// TIA Portal project "session2" (V18)

(* hardware
DEVICE "S7-1200 station_1"  S7-1200 Station
   slot 0: "Rack_0"  S7-1200 Rack  Rack  V1.0
   slot 1: "PLC_1"  CPU 1215C DC/DC/DC  6ES7 215-1AG40-0XB0  V4.6
   slot 2: "SM 1278_1"  4SI IO link  6ES7 278-4BD32-0XB0  V2.1
   slot 3: "DI 2/DQ 2x24VDC_1"  DI2/DQ2 signal board  6ES7 223-0BD30-0XB0  V1.0
DEVICE "HMI_1"  KTP700 Basic PN
   slot 0: "HMI_1"  KTP700 Basic PN  6AV2 123-2GB03-0AX0  17.0.0.0
   slot 1: "HMI_RT_1"  KTP700 Basic PN  6AV2 123-2GB03-0AX0  17.0.0.0
   slot 5: "HMI_1.IE_CP_1"  PROFINET Interface  17.0.0.0
      slot 1: "PROFINET Interface_1"  PROFINET Interface
         slot 1: "Port_1"  Port
DEVICE "GSD device_1"  GSD.Device.PN
   slot 0: "Rack"  Rack  V1.0
   slot 0: "ur3ln"  V1.0  00000
      slot 0: "V1.0"  V1.0
      slot 1: "Interface"  Interface
         slot 1: "RJ45 10/100 MBit/s"  RJ45 10/100 MBit/s
   slot 5: "5_T2O General Purpose Bit Registers_1"  5_T2O General Purpose Bit Registers  1.0
      slot 0: "5_T2O General Purpose Bit Registers"  5_T2O General Purpose Bit Registers
   slot 9: "9_O2T General Purpose Registers 1_1"  9_O2T General Purpose Registers 1  1.0
      slot 0: "9_O2T General Purpose Registers 1"  9_O2T General Purpose Registers 1
*)

// ===== PLC "PLC_1"  CPU 1215C DC/DC/DC =====

VAR_GLOBAL   // PLC tag table "Default tag table"
   "x5" AT %I4.0 : Bool;
   "b1" AT %I1.3 : Bool;
   "b2" AT %I1.4 : Bool;
   "km1" AT %Q1.0 : Bool;
   "km2" AT %Q1.1 : Bool;
   "etap0" AT %M1.0 : Bool;
   "etap1" AT %M1.1 : Bool;
   "etap2" AT %M1.2 : Bool;
   "etap3" AT %M1.3 : Bool;
   "temps" AT %M10.0 : Bool;
   "pos int" AT %MW40 : Word;
   "loop" AT %M12.0 : Bool;
   "input compteur" AT %MW20 : Int;
   "output compteur" AT %MW80 : Int;
   "reset" AT %M5.1 : Bool;
   "Marche" AT %M5.0 : Bool;
   "Temps input" AT %MD30 : Time;
   "temps output" AT %MD34 : Time;
   "Off" AT %M5.2 : Bool;
   "Pos" AT %MW42 : Word;
   "Clock_Byte" AT %MB100 : Byte;
   "Clock_10Hz" AT %M100.0 : Bool;
   "Clock_5Hz" AT %M100.1 : Bool;
   "Clock_2.5Hz" AT %M100.2 : Bool;
   "Clock_2Hz" AT %M100.3 : Bool;
   "Clock_1.25Hz" AT %M100.4 : Bool;
   "Clock_1Hz" AT %M100.5 : Bool;
   "Clock_0.625Hz" AT %M100.6 : Bool;
   "Clock_0.5Hz" AT %M100.7 : Bool;
   "Courant Sig Aut" AT %IW64 : Int;
   "Courant NormX" AT %MD400 : Real;
   "Courant ScaleX" AT %MD500 : Real;
   "Tension Sig Aut" AT %IW66 : Int;
   "Tension NormX" AT %MD600 : Real;
   "Tension ScaleX" AT %MD700 : Real;
   "km4" AT %MW704 : Int;
   "Port Ultrason" AT %IW10 : Word;
   "SubDistance" AT %MW90 : Word;
   "hauteur" AT %MW92 : Word;
   "Distance Manu" AT %MW94 : Word;
   "Nbr Pieces" AT %MW96 : Word;
   "INC" AT %I1.5 : Bool;
   "pos RFID" AT %MW46 : Word;
   "Puc_Data" AT %MW48 : Word;
   "Vitesse" AT %MW110 : Word;
   "Tag_1" AT %QW1000 : Word;
   "Valid" AT %Q150.0 : Bool;
   "Finish" AT %I150.0 : Bool;
   "Err" AT %MW2 : Int;
END_VAR

VAR_GLOBAL   // PLC tag table "RFID_table"
   "RFID_commandBteOut" AT %QB10 : Byte;
   "RFID_CmdStart" AT %Q11.0 : Bool;
   "RFID_CmdDesactivateAntenna" AT %Q11.3 : Bool;
   "RFID_Write_Data1" AT %QW12 : Word;
   "RFID_CommandByteIn" AT %IB10 : Byte;
   "RFID_CmdStartAcknowledge" AT %I11.0 : Bool;
   "RFID_CmdEnd" AT %I11.1 : Bool;
   "RFID_Tag Present" AT %I11.2 : Bool;
   "RFID_Antenna Deactivated" AT %I11.3 : Bool;
   "RFID_Read_Data 1" AT %IW12 : Word;
   "RFID Read_Data2" AT %IW14 : Word;
   "RFID_Read_Data 3" AT %IW16 : Word;
   "RFID_Read_Data4" AT %IW18 : Word;
END_VAR

VAR_GLOBAL   // PLC tag table "Web"
   "Web_CMD_StartMarche" AT %M0.0 : Bool;
   "Web_CMD_StopMarche" AT %M0.1 : Bool;
   "Web_CMD_Reset" AT %M0.2 : Bool;
END_VAR

DATA_BLOCK "Ultrason"   // DB2
{ S7_Optimized_Access := 'TRUE' }
VERSION : 0.1
   VAR
      Distance : Int;
      Hauteur : Int;
      "Nbr Voiture" : Int;
      "Distance 0" : Int := 300;
      inter : Int;
   END_VAR
BEGIN
END_DATA_BLOCK

DATA_BLOCK "Energy Meter"   // DB6
{ S7_Optimized_Access := 'TRUE' }
VERSION : 0.1
   VAR
      Parameter_connexion : TCON_IP_v4;
   END_VAR
BEGIN
   Parameter_connexion.InterfaceId := 64;
   Parameter_connexion.ID := 1;
   Parameter_connexion.ActiveEstablished := true;
   Parameter_connexion.RemoteAddress.ADDR[1] := 172;
   Parameter_connexion.RemoteAddress.ADDR[2] := 28;
   Parameter_connexion.RemoteAddress.ADDR[3] := 111;
   Parameter_connexion.RemoteAddress.ADDR[4] := 56;
   Parameter_connexion.RemotePort := 502;
END_DATA_BLOCK

DATA_BLOCK "node_red"   // DB9
{ S7_Optimized_Access := 'FALSE' }
VERSION : 0.1
   VAR
      courant : Real;
      tension : Real;
   END_VAR
BEGIN
END_DATA_BLOCK

// folder: System blocks/Program resources

DATA_BLOCK "IEC_Timer_0_DB"   // DB1
{ S7_Optimized_Access := 'TRUE' }
AUTHOR : Simatic
FAMILY : IEC
NAME : IEC_TMR
VERSION : 1.0
// stored: InstanceOfName IEC_TIMER
"IEC_TIMER"
BEGIN
END_DATA_BLOCK

DATA_BLOCK "IEC_Counter_0_DB_1"   // DB3
{ S7_Optimized_Access := 'TRUE' }
AUTHOR : Simatic
FAMILY : IEC
NAME : CNTR
VERSION : 1.0
// stored: InstanceOfName IEC_COUNTER
"IEC_COUNTER"
BEGIN
END_DATA_BLOCK

DATA_BLOCK "IEC_Counter_0_DB_2"   // DB4
{ S7_Optimized_Access := 'TRUE' }
AUTHOR : Simatic
FAMILY : IEC
NAME : CNTR
VERSION : 1.0
// stored: InstanceOfName IEC_COUNTER
"IEC_COUNTER"
BEGIN
END_DATA_BLOCK

DATA_BLOCK "IEC_Counter_0_DB"   // DB7
{ S7_Optimized_Access := 'TRUE' }
AUTHOR : Simatic
FAMILY : IEC
NAME : CNTR
VERSION : 1.0
// stored: InstanceOfName IEC_COUNTER
"IEC_COUNTER"
BEGIN
END_DATA_BLOCK

// folder: (top level)

FUNCTION "configurer" : Void   // FC1, LAD
{ S7_Optimized_Access := 'TRUE' }
VERSION : 0.1
BEGIN

REGION Network 1
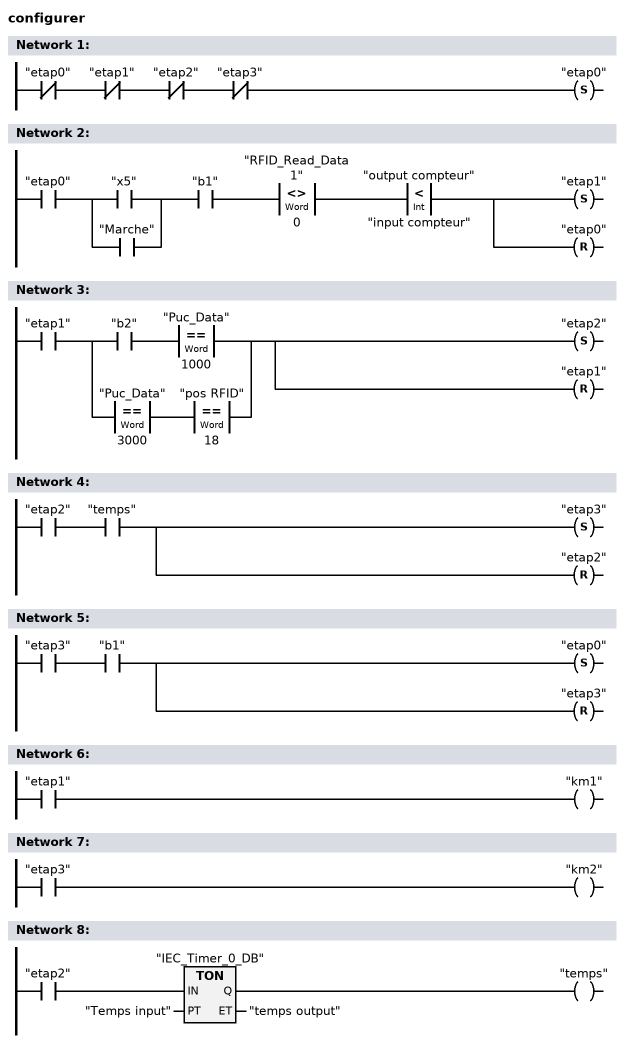
   RUNG wire#powerrail
      I_Contact( "etap0" )
      I_Contact( "etap1" )
      I_Contact( "etap2" )
      I_Contact( "etap3" )
      S_Coil( "etap0" )
   END_RUNG
   // the same network as SCL:
   IF NOT "etap0" AND NOT "etap1" AND NOT "etap2" AND NOT "etap3" THEN "etap0" := TRUE; END_IF;
END_REGION

REGION Network 2
   RUNG wire#powerrail
      Contact( "etap0" )
      wire#w1
      Contact( "x5" )
      wire#w2
      Contact( "b1" )
      { S7_Templates := "SrcType := Word" } NE_Contact(in1 := "RFID_Read_Data 1", in2 := 0)
      { S7_Templates := "SrcType := Int" } LT_Contact(in1 := "output compteur", in2 := "input compteur")
      wire#w3
      S_Coil( "etap1" )
   END_RUNG
   RUNG wire#w1
      Contact( "Marche" )
   END_RUNG wire#w2
   RUNG wire#w3
      R_Coil( "etap0" )
   END_RUNG
   // the same network as SCL:
   IF "etap0" AND ("x5" OR "Marche") AND "b1" AND ("RFID_Read_Data 1" <> 0) AND ("output compteur" < "input compteur") THEN
       "etap1" := TRUE;
       "etap0" := FALSE;
   END_IF;
END_REGION

REGION Network 3
   RUNG wire#powerrail
      Contact( "etap1" )
      wire#w1
      Contact( "b2" )
      { S7_Templates := "SrcType := Word" } EQ_Contact(in1 := "Puc_Data", in2 := 1000)
      wire#w2
      S_Coil( "etap2" )
   END_RUNG
   RUNG wire#w1
      { S7_Templates := "SrcType := Word" } EQ_Contact(in1 := "Puc_Data", in2 := 3000)
      { S7_Templates := "SrcType := Word" } EQ_Contact(in1 := "pos RFID", in2 := 18)
   END_RUNG wire#w2
   RUNG wire#w2
      R_Coil( "etap1" )
   END_RUNG
   // the same network as SCL:
   IF "etap1" AND (("b2" AND ("Puc_Data" = 1000)) OR (("Puc_Data" = 3000) AND ("pos RFID" = 18))) THEN
       "etap2" := TRUE;
       "etap1" := FALSE;
   END_IF;
END_REGION

REGION Network 4
   RUNG wire#powerrail
      Contact( "etap2" )
      Contact( "temps" )
      wire#w1
      S_Coil( "etap3" )
   END_RUNG
   RUNG wire#w1
      R_Coil( "etap2" )
   END_RUNG
   // the same network as SCL:
   IF "etap2" AND "temps" THEN
       "etap3" := TRUE;
       "etap2" := FALSE;
   END_IF;
END_REGION

REGION Network 5
   RUNG wire#powerrail
      Contact( "etap3" )
      Contact( "b1" )
      wire#w1
      S_Coil( "etap0" )
   END_RUNG
   RUNG wire#w1
      R_Coil( "etap3" )
   END_RUNG
   // the same network as SCL:
   IF "etap3" AND "b1" THEN
       "etap0" := TRUE;
       "etap3" := FALSE;
   END_IF;
END_REGION

REGION Network 6
   RUNG wire#powerrail
      Contact( "etap1" )
      Coil( "km1" )
   END_RUNG
   // the same network as SCL:
   "km1" := "etap1";
END_REGION

REGION Network 7
   RUNG wire#powerrail
      Contact( "etap3" )
      Coil( "km2" )
   END_RUNG
   // the same network as SCL:
   "km2" := "etap3";
END_REGION

REGION Network 8
   "IEC_Timer_0_DB".TON(IN := "etap2", PT := "Temps input", ET => "temps output");
   "temps" := "IEC_Timer_0_DB".Q;
END_REGION
END_FUNCTION

FUNCTION "Conversion" : Void   // FC2, LAD
{ S7_Optimized_Access := 'TRUE' }
VERSION : 0.1
BEGIN

REGION Network 1
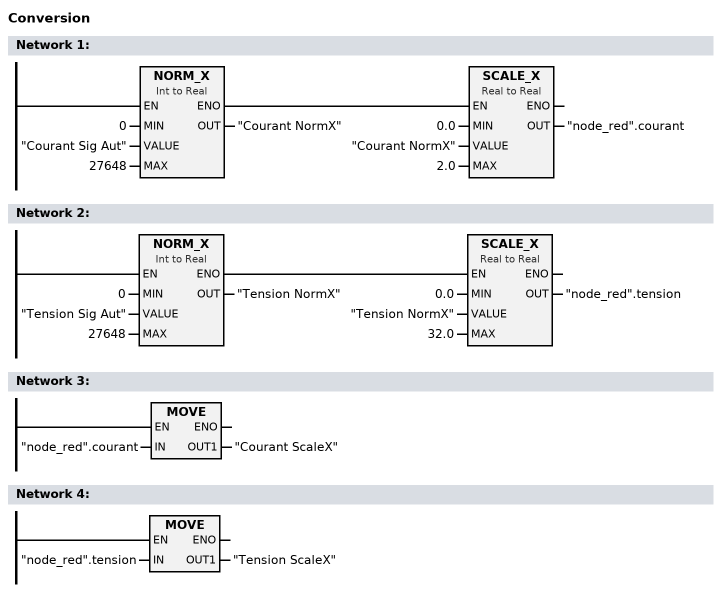
   RUNG wire#powerrail
      { S7_Templates := "[SrcType := Int, DestType := Real]" } Normalize(min := 0, value := "Courant Sig Aut", max := 27648, out => "Courant NormX")
      { S7_Templates := "[SrcType := Real, DestType := Real]" } Scale(min := 0.0, value := "Courant NormX", max := 2.0, out => "node_red".courant)
   END_RUNG
   // the same network as SCL:
   "Courant NormX" := NORM_X(MIN := 0, VALUE := "Courant Sig Aut", MAX := 27648);
   "node_red".courant := SCALE_X(MIN := 0.0, VALUE := "Courant NormX", MAX := 2.0);
END_REGION

REGION Network 2
   RUNG wire#powerrail
      { S7_Templates := "[SrcType := Int, DestType := Real]" } Normalize(min := 0, value := "Tension Sig Aut", max := 27648, out => "Tension NormX")
      { S7_Templates := "[SrcType := Real, DestType := Real]" } Scale(min := 0.0, value := "Tension NormX", max := 32.0, out => "node_red".tension)
   END_RUNG
   // the same network as SCL:
   "Tension NormX" := NORM_X(MIN := 0, VALUE := "Tension Sig Aut", MAX := 27648);
   "node_red".tension := SCALE_X(MIN := 0.0, VALUE := "Tension NormX", MAX := 32.0);
END_REGION

REGION Network 3
   RUNG wire#powerrail
      Move(in := "node_red".courant, out1 => "Courant ScaleX")
   END_RUNG
   // the same network as SCL:
   "Courant ScaleX" := "node_red".courant;
END_REGION

REGION Network 4
   RUNG wire#powerrail
      Move(in := "node_red".tension, out1 => "Tension ScaleX")
   END_RUNG
   // the same network as SCL:
   "Tension ScaleX" := "node_red".tension;
END_REGION
END_FUNCTION

FUNCTION "Ultrason Configuration" : Void   // FC3, LAD
{ S7_Optimized_Access := 'TRUE' }
VERSION : 0.1
   VAR_TEMP
      "inter 1" : Int;
   END_VAR
BEGIN

REGION Network 1
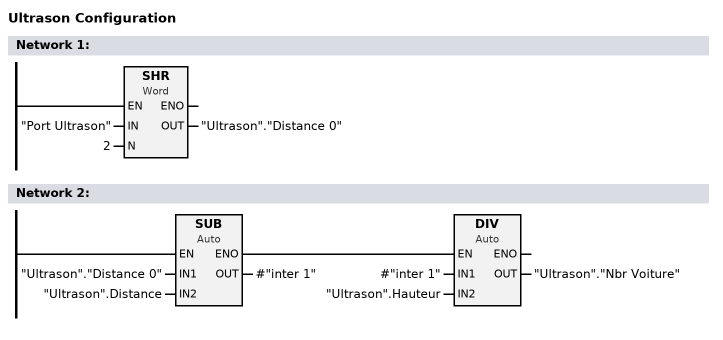
   RUNG wire#powerrail
      { S7_Templates := "SrcType := Word" } Shr(in := "Port Ultrason", n := 2, out => "Ultrason"."Distance 0")
   END_RUNG
   // the same network as SCL:
   "Ultrason"."Distance 0" := SHR(IN := "Port Ultrason", N := 2);
END_REGION

REGION Network 2
   RUNG wire#powerrail
      Sub(in1 := "Ultrason"."Distance 0", in2 := "Ultrason".Distance, out => #"inter 1")
      Div(in1 := #"inter 1", in2 := "Ultrason".Hauteur, out => "Ultrason"."Nbr Voiture")
   END_RUNG
   // the same network as SCL:
   #"inter 1" := "Ultrason"."Distance 0" - "Ultrason".Distance;
   "Ultrason"."Nbr Voiture" := #"inter 1" / "Ultrason".Hauteur;
END_REGION
END_FUNCTION

FUNCTION "Central de Mesure" : Void   // FC4, LAD
{ S7_Optimized_Access := 'TRUE' }
VERSION : 0.1
BEGIN

REGION Network 1
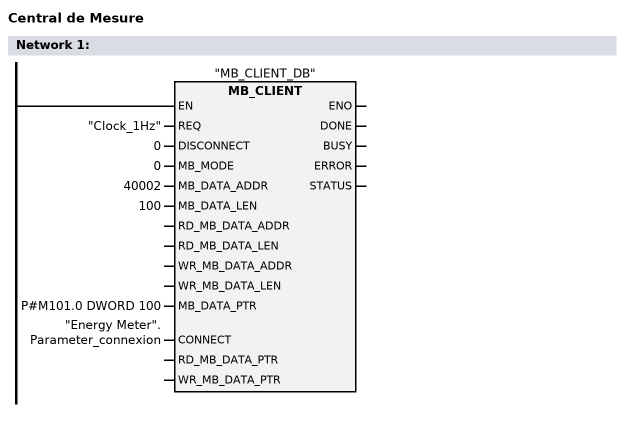
   "MB_CLIENT_DB"(REQ := "Clock_1Hz",   // MB_CLIENT
                  DISCONNECT := 0,
                  MB_MODE := 0,
                  MB_DATA_ADDR := 40002,
                  MB_DATA_LEN := 100,
                  MB_DATA_PTR := P#M101.0 DWORD 100,
                  CONNECT := "Energy Meter".Parameter_connexion);
END_REGION
END_FUNCTION

FUNCTION "WebServerTesting" : Void   // FC5, LAD
{ S7_Optimized_Access := 'TRUE' }
VERSION : 0.1
BEGIN

REGION Network 1
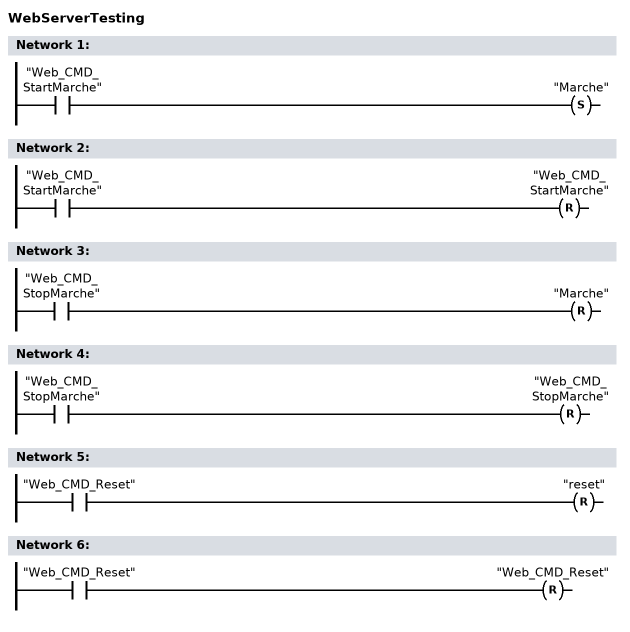
   RUNG wire#powerrail
      Contact( "Web_CMD_StartMarche" )
      S_Coil( "Marche" )
   END_RUNG
   // the same network as SCL:
   IF "Web_CMD_StartMarche" THEN "Marche" := TRUE; END_IF;
END_REGION

REGION Network 2
   RUNG wire#powerrail
      Contact( "Web_CMD_StartMarche" )
      R_Coil( "Web_CMD_StartMarche" )
   END_RUNG
   // the same network as SCL:
   IF "Web_CMD_StartMarche" THEN "Web_CMD_StartMarche" := FALSE; END_IF;
END_REGION

REGION Network 3
   RUNG wire#powerrail
      Contact( "Web_CMD_StopMarche" )
      R_Coil( "Marche" )
   END_RUNG
   // the same network as SCL:
   IF "Web_CMD_StopMarche" THEN "Marche" := FALSE; END_IF;
END_REGION

REGION Network 4
   RUNG wire#powerrail
      Contact( "Web_CMD_StopMarche" )
      R_Coil( "Web_CMD_StopMarche" )
   END_RUNG
   // the same network as SCL:
   IF "Web_CMD_StopMarche" THEN "Web_CMD_StopMarche" := FALSE; END_IF;
END_REGION

REGION Network 5
   RUNG wire#powerrail
      Contact( "Web_CMD_Reset" )
      R_Coil( "reset" )
   END_RUNG
   // the same network as SCL:
   IF "Web_CMD_Reset" THEN "reset" := FALSE; END_IF;
END_REGION

REGION Network 6
   RUNG wire#powerrail
      Contact( "Web_CMD_Reset" )
      R_Coil( "Web_CMD_Reset" )
   END_RUNG
   // the same network as SCL:
   IF "Web_CMD_Reset" THEN "Web_CMD_Reset" := FALSE; END_IF;
END_REGION
END_FUNCTION

ORGANIZATION_BLOCK "Main"   // OB1, LAD, ProgramCycle
{ S7_Optimized_Access := 'TRUE' }
VERSION : 0.1
   VAR_INPUT
      Initial_Call : Bool;
      Remanence : Bool;
   END_VAR
BEGIN

REGION Network 1
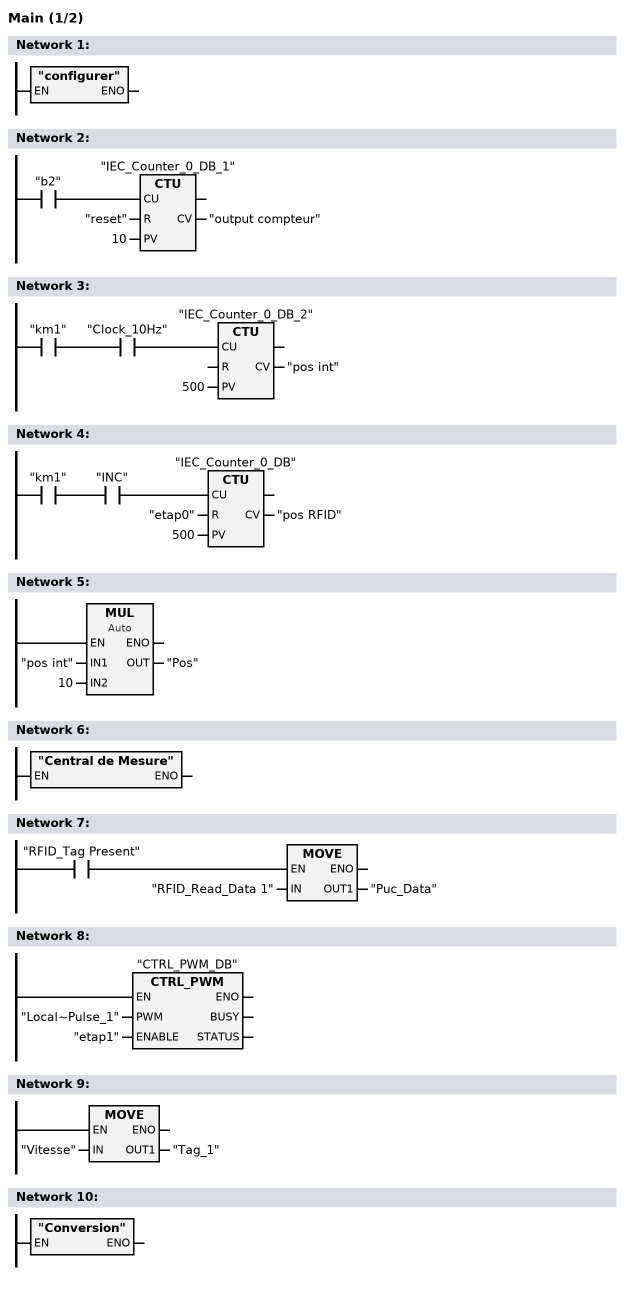
   RUNG wire#powerrail
      "configurer"()
   END_RUNG
   // the same network as SCL:
   "configurer"();
END_REGION

REGION Network 2
   "IEC_Counter_0_DB_1".CTU(CU := "b2", R := "reset", PV := 10, CV => "output compteur");
END_REGION

REGION Network 3
   "IEC_Counter_0_DB_2".CTU(CU := "km1" AND "Clock_10Hz", PV := 500, CV => "pos int");
END_REGION

REGION Network 4
   "IEC_Counter_0_DB".CTU(CU := "km1" AND "INC", R := "etap0", PV := 500, CV => "pos RFID");
END_REGION

REGION Network 5
   RUNG wire#powerrail
      Mul(in1 := "pos int", in2 := 10, out => "Pos")
   END_RUNG
   // the same network as SCL:
   "Pos" := "pos int" * 10;
END_REGION

REGION Network 6
   RUNG wire#powerrail
      "Central de Mesure"()
   END_RUNG
   // the same network as SCL:
   "Central de Mesure"();
END_REGION

REGION Network 7
   RUNG wire#powerrail
      Contact( "RFID_Tag Present" )
      Move(in := "RFID_Read_Data 1", out1 => "Puc_Data")
   END_RUNG
   // the same network as SCL:
   IF "RFID_Tag Present" THEN "Puc_Data" := "RFID_Read_Data 1"; END_IF;
END_REGION

REGION Network 8
   "CTRL_PWM_DB"(PWM := "Local~Pulse_1", ENABLE := "etap1");   // CTRL_PWM
END_REGION

REGION Network 9
   RUNG wire#powerrail
      Move(in := "Vitesse", out1 => "Tag_1")
   END_RUNG
   // the same network as SCL:
   "Tag_1" := "Vitesse";
END_REGION

REGION Network 10
   RUNG wire#powerrail
      "Conversion"()
   END_RUNG
   // the same network as SCL:
   "Conversion"();
END_REGION

REGION Network 11
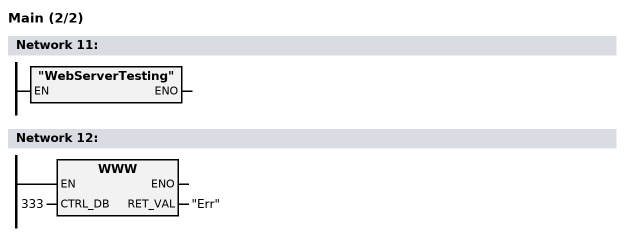
   RUNG wire#powerrail
      "WebServerTesting"()
   END_RUNG
   // the same network as SCL:
   "WebServerTesting"();
END_REGION

REGION Network 12
   "Err" := WWW(CTRL_DB := 333);
END_REGION
END_ORGANIZATION_BLOCK

(* ===== HMI "HMI_RT_1" =====
system functions are stored by id; their names below are inferred from use
connection "HMI_Connection_1": ETHERNET, SMART_S7_1200_OMS

HMI tags "Default tag table"
   "Tag_ScreenNumber" : UInt, internal
   "b1" : Bool = PLC b1 AT %I1.3, 1 s
   "b2" : Bool = PLC b2 AT %I1.4, 1 s
   "output compteur" : Int = PLC "output compteur" AT %MW80, 1 s
   "reset" : Bool = PLC reset AT %M5.1, 1 s
   "Tag_1" : Bool = PLC Marche AT %M5.0, 1 s
   "input compteur" : Int = PLC "input compteur" AT %MW20, 1 s
   "Temps input" : Time = PLC "Temps input" AT %MD30, 1 s
   "temps output" : Time = PLC "temps output" AT %MD34, 1 s
   "Off" : Bool = PLC Off AT %M5.2, 1 s
   "km1" : Bool = PLC km1 AT %Q1.0, 1 s
   "km2" : Bool = PLC km2 AT %Q1.1, 1 s
   "Pos(1)" : Word = PLC Pos AT %MW42, 1 s
   "Courant ScaleX" : Real = PLC "Courant ScaleX" AT %MD500, 1 s
   "Tension ScaleX" : Real = PLC "Tension ScaleX" AT %MD700, 1 s
   "Distance Manu" : Word = PLC "Distance Manu" AT %MW94, 1 s
   "hauteur" : Word = PLC hauteur AT %MW92, 1 s
   "Nbr Pieces" : Word = PLC "Nbr Pieces" AT %MW96, 1 s
   "Ultrason_Distance 0" : Int = PLC Ultrason."Distance 0", 1 s
   "Ultrason_Hauteur" : Int = PLC Ultrason.Hauteur, 1 s
   "Ultrason_Nbr Voiture" : Int = PLC Ultrason."Nbr Voiture", 1 s
   "Ultrason_Distance" : Int = PLC Ultrason.Distance, 1 s
   "RFID_commandBteOut" : Byte = PLC RFID_commandBteOut AT %QB10, 1 s
   "RFID_Write_Data1" : Word = PLC RFID_Write_Data1 AT %QW12, 1 s
   "RFID_CmdStart" : Bool = PLC RFID_CmdStart AT %Q11.0, 1 s
   "RFID_Antenna Deactivated" : Bool = PLC "RFID_Antenna Deactivated" AT %I11.3, 1 s
   "RFID_Read_Data 1" : Word = PLC "RFID_Read_Data 1" AT %IW12, 1 s
   "RFID_Tag Present" : Bool = PLC "RFID_Tag Present" AT %I11.2, 1 s
   "RFID_CmdEnd" : Bool = PLC RFID_CmdEnd AT %I11.1, 1 s
   "pos RFID" : Word = PLC "pos RFID" AT %MW46, 1 s
   "Vitesse" : Word = PLC Vitesse AT %MW110, 1 s

Template "Tunisia" 800x480
   SymbolicIOField "Symbolic_IO_Field_Screen" at 93,9 size 600x33; TextOff '0'; TextOn '1'; TextList "TextList_ScreenNames"
      ProcessValue <- "Tag_ScreenNumber"
      on Change: ActivateScreenByNumber("Tag_ScreenNumber", 0)
   DateTimeField "HmiScreenItemData" at 695,25 size 105x25
   DateTimeField "HmiScreenItemData_1" at 695,0 size 105x25
   GraphicView "Graphic view_3" at 701,8 size 73x36; Picture "Graphic_6"

screen "Root screen" 800x480, template "Tunisia"
   on GenerateScreen: SetTag("Tag_ScreenNumber", 1)
   TextField "HmiScreenItemData_1" at 64,435 size 640x25; Text 'Welcome User !!'
   Button "HmiScreenItemData" at 163,124 size 159x47; TextOff 'convoyer'; PictureOff "Navigates to convoyer for KTP700 Basic+ PN 17.0.0.0"; PictureOn "Navigates to convoyer for KTP700 Basic+ PN 17.0.0.0"
      on Release: ActivateScreen("convoyer", 0)
   Button "HmiScreenItemData_2" at 163,296 size 159x47; TextOn 'convoyer'; TextOff 'Mesure Ultrason'; PictureOn "Navigates to convoyer for KTP700 Basic+ PN 17.0.0.0"; PictureOff "Navigates to convoyer for KTP700 Basic+ PN 17.0.0.0"
      on Release: ActivateScreen("Mesure Ultrason", 0)
   Button "HmiScreenItemData_3" at 163,180 size 159x47; TextOn 'convoyer'; TextOff 'RFID'; PictureOn "Navigates to convoyer for KTP700 Basic+ PN 17.0.0.0"; PictureOff "Navigates to convoyer for KTP700 Basic+ PN 17.0.0.0"
      on Release: ActivateScreen("RFID", 0)
   Button "HmiScreenItemData_4" at 163,238 size 159x47; TextOn 'convoyer'; TextOff 'Position'; PictureOn "Navigates to convoyer for KTP700 Basic+ PN 17.0.0.0"; PictureOff "Navigates to convoyer for KTP700 Basic+ PN 17.0.0.0"
      on Release: ActivateScreen("Position", 0)
   GraphicView "Graphic view_1" at 286,425 size 36x30; Picture "Graphic_5"
   GraphicView "Graphic view_2" at 379,167 size 201x134; Picture "Graphic_6"

screen "convoyer" 800x480, template "Tunisia"
   on GenerateScreen: SetTag("Tag_ScreenNumber", 2)
   TextField "HmiScreenItemData" at 307,262 size 165x25; Text 'convoyer'
   Button "Back" at 666,423 size 109x37; TextOff 'Back'
      on Release: ActivateScreen("Root screen", 0)
   Circle "Circle_1" at 260,213 size 48x48
      Appearance <- "km1"
   Circle "Circle_2" at 487,213 size 48x48
      Appearance <- "km2"
   Rectangle "Rectangle_1" at 277,214 size 15x46
      Appearance <- "b1"
   Rectangle "Rectangle_2" at 505,213 size 15x46
      Appearance <- "b2"
   Button "Button_1" at 671,164 size 96x32; TextOff 'Reset'
      on Press: SetBit("reset")
      on Release: ResetBit("reset")
   IOField "I/O field_1" at 450,119 size 102x32; FormatPattern 999; Unit  Piéces
      ProcessValue <- "output compteur"
   TextField "Text field_1" at 268,121 size 181x23; Text 'Valeur du compteur :'
   Button "Button_2" at 670,118 size 96x32; TextOff 'Off'
      on Press: ResetBit("Tag_1")
   Button "Button_3" at 670,76 size 96x32; TextOff 'On'
      on Press: SetBit("Tag_1")
   IOField "I/O field_2" at 449,72 size 102x32; FormatPattern 999; Unit  Piéces
      ProcessValue <- "input compteur"
   TextField "Text field_2" at 268,74 size 175x23; Text 'Nombre des Piéces :'
   IOField "I/O field_3" at 450,370 size 102x32; FormatPattern 9999; Unit  ms
      ProcessValue <- "temps output"
   TextField "Text field_3" at 268,372 size 128x23; Text 'Temps Ecoulé :'
   IOField "I/O field_4" at 449,325 size 102x32; FormatPattern 9999; Unit  ms
      ProcessValue <- "Temps input"
   TextField "Text field_4" at 268,325 size 116x23; Text 'Fixer Temps :'
   GraphicView "Graphic view_1" at 34,93 size 95x75; Picture "Graphic_7"
      Visibility <- "km1"
   GraphicView "Graphic view_2" at 34,201 size 95x75; Picture "Graphic_8"
      Visibility <- "km2"
   Rectangle "Rectangle_10" at 287,191 size 30x23
      HorizontalMovement <- "Pos(1)"
   TextField "Text field_5" at 31,62 size 101x23; Text 'Moteur On :'
   TextField "Text field_6" at 27,173 size 83x23; Text 'Moteur 1'
   TextField "Text field_7" at 29,279 size 83x23; Text 'Moteur 2'
   IOField "I/O field_5" at 35,325 size 96x32; FormatPattern 99.999; Unit  A
      ProcessValue <- "Courant ScaleX"
   IOField "I/O field_6" at 36,372 size 96x32; FormatPattern 99.999; Unit  V
      ProcessValue <- "Tension ScaleX"
   TextField "Text field_8" at 36,307 size 66x20; Text 'Courant :'
   TextField "Text field_9" at 36,354 size 63x20; Text 'Tension :'
   IOField "I/O field_7" at 671,240 size 96x32; FormatPattern 99999
      ProcessValue <- "pos RFID"
   TextField "Text field_10" at 678,210 size 71x23; Text 'Position'
   IOField "I/O field_8" at 671,302 size 96x32; FormatPattern 99999
      ProcessValue <- "Vitesse"
   TextField "Text field_11" at 678,276 size 64x23; Text 'Vitesse'
   GraphicView "Graphic view_3" at 34,93 size 95x75; Picture "Graphic_10"
      Visibility <- "km1"
   GraphicView "Graphic view_4" at 34,201 size 95x75; Picture "Graphic_10"
      Visibility <- "km2"

screen "RFID" 800x480, template "Tunisia"
   TextField "Text field_1" at 174,58 size 67x27; Text 'INPUT'
   TextField "Text field_2" at 546,58 size 84x27; Text 'OUTPUT'
   Button "Button_1" at 440,106 size 292x32; TextOff 'Read'
      on Press: SetTag("RFID_commandBteOut", 1)
      Appearance <- "RFID_commandBteOut"
   Button "Button_3" at 444,170 size 292x32; TextOff 'Write'
      on Press: SetTag("RFID_commandBteOut", 2)
      Appearance <- "RFID_commandBteOut"
   Button "Button_2" at 440,387 size 292x32; TextOff 'Start'
      on Press: function_b14e0dd5("RFID_CmdStart", 0)
   IOField "I/O field_1" at 440,323 size 85x34; FormatPattern 99999
      ProcessValue <- "RFID_Write_Data1"
   TextField "Text field_3" at 577,325 size 131x27; Text 'Data to write'
   Rectangle "Rectangle_5" at 82,106 size 253x51
      Appearance <- "RFID_Antenna Deactivated"
   Rectangle "Rectangle_6" at 82,170 size 253x51
      Appearance <- "RFID_Tag Present"
   Rectangle "Rectangle_7" at 82,232 size 253x51
      Appearance <- "RFID_CmdStart"
   Rectangle "Rectangle_8" at 82,295 size 253x51
      Appearance <- "RFID_CmdEnd"
   IOField "I/O field_2" at 256,372 size 85x34; FormatPattern 99999
      ProcessValue <- "RFID_Read_Data 1"
   TextField "Text field_4" at 103,375 size 123x27; Text 'Data to read'
   TextField "Text field_8" at 137,115 size 143x32; Text 'Antenna off'
      Visibility <- "RFID_Antenna Deactivated"
   TextField "Text field_5" at 155,305 size 108x32; Text 'CMD End'
   TextField "Text field_6" at 132,241 size 152x32; Text 'CMD Started'
   TextField "Text field_7" at 136,179 size 144x32; Text 'Tag Present'
   TextField "Text field_9" at 137,115 size 140x32; Text 'Antenna on'
      Visibility <- "RFID_Antenna Deactivated"
   Button "Back" at 86,418 size 109x37; TextOn 'Back'; TextOff 'Back'
      on Release: ActivateScreen("Root screen", 0)
   IOField "I/O field_3" at 546,241 size 96x32; FormatPattern 99999
      ProcessValue <- "pos RFID"
   TextField "Text field_10" at 553,211 size 71x23; Text 'Position'

screen "Mesure Ultrason" 800x480, template "Tunisia"
   IOField "I/O field_1" at 62,109 size 97x32; FormatPattern 9999; Unit  cm
      ProcessValue <- "Ultrason_Distance 0"
   IOField "I/O field_2" at 62,230 size 98x32; FormatPattern 9999; Unit  cm
      ProcessValue <- "Ultrason_Hauteur"
   IOField "I/O field_3" at 54,404 size 112x32; FormatPattern 9999; Unit  piéces
      ProcessValue <- "Ultrason_Nbr Voiture"
   TextField "Text field_1" at 71,86 size 90x23; Text 'Distance 0'
   TextField "Text field_2" at 71,207 size 71x23; Text 'Hauteur'
   TextField "Text field_3" at 39,379 size 140x23; Text 'Nbr des Voitures'
   GraphicView "Graphic view_1" at 62,309 size 105x57; Picture "Graphic_2"
   Button "Back" at 666,423 size 109x37; TextOn 'Back'; TextOff 'Back'
      on Release: ActivateScreen("Root screen", 0)
   IOField "I/O field_4" at 61,167 size 97x32; FormatPattern 9999; Unit  cm
      ProcessValue <- "Ultrason_Distance"
   TextField "Text field_4" at 70,144 size 75x23; Text 'Distance'
   GraphicView "Graphic view_2" at 433,120 size 89x102; Picture "images"

screen "Position" 800x480, template "Tunisia"
   Button "Back" at 86,398 size 109x37; TextOn 'Back'; TextOff 'Back'
      on Release: ActivateScreen("Root screen", 0)
   IOField "I/O field_1" at 357,191 size 96x32; FormatPattern 99999
      ProcessValue <- "pos RFID"
   TextField "Text field_1" at 364,161 size 71x23; Text 'Position'
*)